(* PLC project c.project, CODESYS CODESYS V3.5 SP17 Patch 3 *)
(* stored: creationDateTime 2026-10-19T00:00:00, modificationDateTime 2026-10-19T00:00:00 *)

FUNCTION_BLOCK FB_C
VAR_INPUT
    i1 : INT;
    i2 : INT;
    s : BOOL;
END_VAR
VAR_OUTPUT
    o : INT;
END_VAR

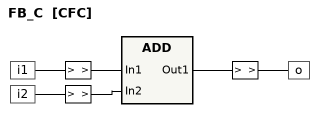
(* CFC diagram, written out as Structured Text *)
o := i1 + i2;
END_FUNCTION_BLOCK
